(* IEC 61131-3 sources: codesys-to-astra/src/POUs/F_C2aAfter, 2 files *)

(* ---- F_C2aAfter.decl.st ---- *)
// Назначение: замена OSU.After (OwenStringUtils v3.0, с. 19): фрагмент sSource после первого вхождения
//             sPrefix; не найдено — пустая строка.
// Автор:      kr0nsch
// Версия:     0.1.0
// Документ:   docs/LIBMAP.md
FUNCTION F_C2aAfter : STRING(255)
VAR_INPUT
    sSource : STRING(255);  // исходная строка
    sPrefix : STRING(255);  // подстрока
END_VAR
VAR
    iPos : INT;             // позиция вхождения (с 1) или 0
END_VAR

(* ---- F_C2aAfter.impl.st ---- *)
iPos := FIND(sSource, sPrefix);
IF iPos > 0 AND LEN(sPrefix) > 0 THEN
    F_C2aAfter := RIGHT(sSource, LEN(sSource) - iPos - LEN(sPrefix) + 1);
ELSE
    F_C2aAfter := '';
END_IF
